VISUALIZATION teste  // 1024x768
END_VISUALIZATION

(* stored: Version 1.1.0.1
   Visu teste: Id {35f59e62-3a7f-4d1f-851a-9c2954d1b78a} *)
